Fanuc KAREL source: KT00234.KL

PROGRAM KT00234
%NOLOCKGROUP
VAR
  I1: INTEGER
  B2: BOOLEAN
  OUT: INTEGER
BEGIN
  I1 = 2
    B2 = FALSE
  OUT = I1 OR B2
END KT00234
